(* Logix 5000 project; controller Soda_Pop_Machine 5069-L306ERM rev 38.11; software revision 38.02 *)

TASK MainTask (continuous, watchdog 500 ms) : MainProgram

MODULES
   Local : 5069-L306ERM (5069 0, rev 38.11)
       : 5069-IB16 (5069 1, rev 2.16, StandardDataDriven RPI 5 ms)
       : 5069-OB16 (5069 2, rev 3.13, StandardDataDriven RPI 5 ms)
       : 5069-IF8 (5069 3, rev 3.11, StandardDataDriven RPI 100 ms)
       : vendor 1 type 115 code 320 (5069 4, rev 2.13, StandardDataDriven RPI 80 ms)
END_MODULES

PROGRAM MainProgram   (* main routine Main *)
VAR
   Add_ice : SFC_STEP := (Status := 16#0020_0001, PauseTimer := 1, PRE := 3000);
   Add_ice_action : SFC_ACTION := (Status := 16#0020_0000, PauseTimer := 1);
   Coin : BOOL;
   Cup : STRING;
   DISPENSE : SFC_STEP := (Status := 16#0020_0001, PauseTimer := 1, PRE := 2000);
   Dispense_action : SFC_ACTION := (Status := 16#0020_0000, PauseTimer := 1);
   Drop_Cup : SFC_STEP := (Status := 16#0020_0001, PauseTimer := 1);
   Enter : BOOL;
   Finish : SFC_STEP := (Status := 16#0020_0001, PauseTimer := 1);
   Flash_lights : SFC_ACTION := (Status := 16#0020_0000, PauseTimer := 1);
   GrapeSTR : STRING := 'Grape';
   IceSTR : STRING := ' + Ice';
   INIT : SFC_STEP := (Status := 16#a820_0201, X := 1, SA := 1, DN := 1, PauseTimer := 1, T := 18659, TMax := 18659, Count := 1);
   Init_action : SFC_ACTION := (Status := 16#c020_0000, A := 1, Q := 1, PauseTimer := 1, Count := 1);
   LED_1 : ALIAS FOR Local:2:O.Pt00.Data;
   LED_2 : ALIAS FOR Local:2:O.Pt01.Data;
   LemonSTR : STRING := 'Lemon';
   Mixer_on : SFC_STEP := (Status := 16#0020_0001, PauseTimer := 1);
   Music_on : SFC_STEP := (Status := 16#0020_0001, PauseTimer := 1);
   Music_on_action : SFC_ACTION := (Status := 16#0020_0000, PauseTimer := 1);
   NullSTR : STRING;
   OrangeSTR : STRING := 'Orange';
   Pass_to_finish : BOOL;
   Pass_to_mixer : BOOL;
   Pass_to_mixer_action : SFC_ACTION := (Status := 16#0020_0000, PauseTimer := 1);
   PeachSTR : STRING := 'Peach';
   pop_type : STRING;
   Return_to_init : BOOL;
   SELECT : SFC_STEP := (Status := 16#0020_0001, PauseTimer := 1);
   Select_action : SFC_ACTION := (Status := 16#0020_0000, PauseTimer := 1);
   Socket_1 : ALIAS FOR Local:2:O.Pt02.Data;
   Socket_2 : ALIAS FOR Local:2:O.Pt03.Data;
   Switch_1 : ALIAS FOR Local:1:I.Pt00.Data;
   Switch_2 : ALIAS FOR Local:1:I.Pt01.Data;
   Switch_3 : ALIAS FOR Local:1:I.Pt02.Data;
   Switch_4 : ALIAS FOR Local:1:I.Pt03.Data;
   Switch_5 : ALIAS FOR Local:1:I.Pt04.Data;
   Switch_6 : ALIAS FOR Local:1:I.Pt05.Data;
   Wait_for_drop : BOOL;
   Wait_for_mixer : BOOL;
   Wait_for_mixer_action : SFC_ACTION := (Status := 16#0020_0000, PauseTimer := 1);
END_VAR

ROUTINE Main   (* sequential function chart *)
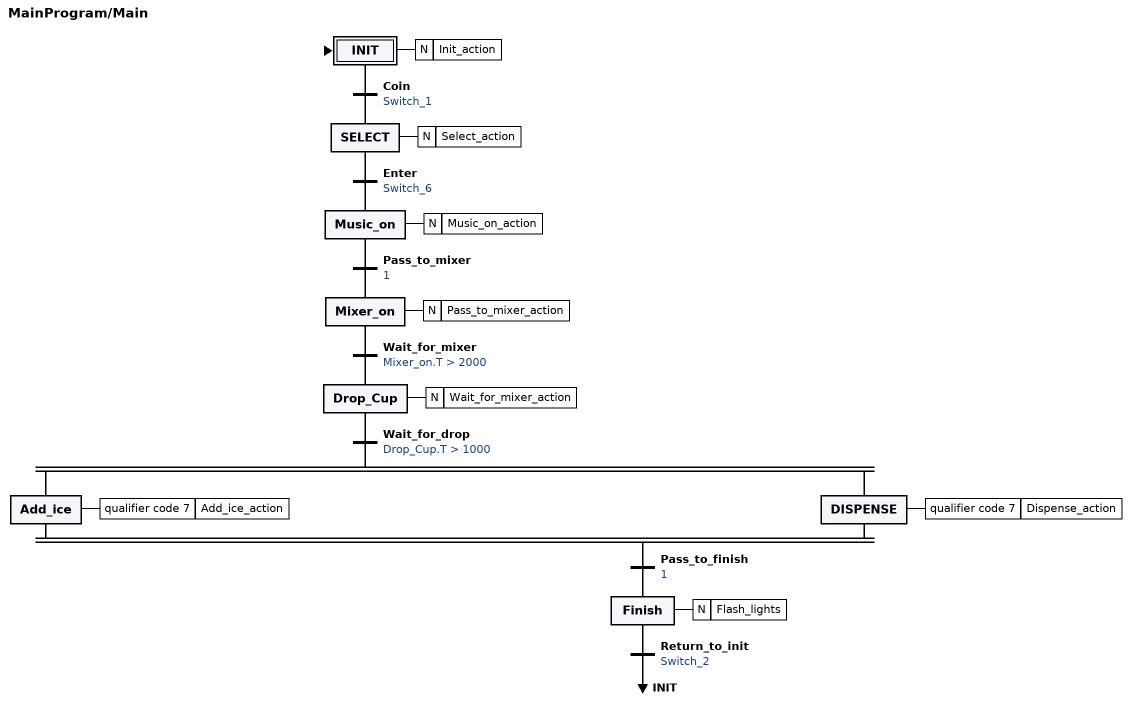
   // "add_ice"
   // step has a
   // preset wait
   // time of 3
   // seconds
   // (3000 ms)
   // "DISPENSE" step
   // has a preset wait
   // time of 2 seconds
   // (2000 ms)
   // Set initial values.
   // Turn off all LEDs
   // and sockets
   // (LEDs 3 and 4).
   // Erase cup string.
   // Select stage
   // represents the
   // customer
   // selecting a
   // options. Turn on
   // LED1 and flash
   // LED2 at 1 Hz.
   // Turn on the
   // music
   // (socket_1,
   // which is actually
   // LED3)
   // Turn on the
   // mixer (socket_2,
   // which is
   // actually LED4)
   // Wait for the
   // mixer for two
   // seconds before
   // continuing.
   // Turn off the
   // mixer. (Turn off
   // Socket_2, LED4)
   // Change the pop
   // type in the "cup"
   // string based off
   // switches 4 and
   // 5.
   // Display a
   // cascading
   // effect of LEDs
   // when finished.
   // Wait for switch
   // 2 before
   // resetting the
   // machine.
   // Wait for for the
   // selections to be
   // entered (switch
   // 6) before
   // continuing.
   INITIAL_STEP INIT:
      ACTION Init_action (N):
         LED_1 := 0;
         LED_2 := 0;
         Socket_1 := 0;
         Socket_2 := 0;
         CONCAT(NullSTR, NullSTR, Cup);
         
      END_ACTION
   END_STEP
   TRANSITION Coin FROM INIT TO SELECT
      := Switch_1
   END_TRANSITION
   STEP SELECT:
      ACTION Select_action (N):
         LED_1 := 1;
         LED_2 := ((SELECT.T / 500) MOD 2) = 0;
         
      END_ACTION
   END_STEP
   TRANSITION Enter FROM SELECT TO Music_on
      := Switch_6
   END_TRANSITION
   STEP Music_on:
      ACTION Music_on_action (N):
         Socket_1 := 1;
      END_ACTION
   END_STEP
   TRANSITION Pass_to_mixer FROM Music_on TO Mixer_on
      := 1
         
   END_TRANSITION
   STEP Mixer_on:
      ACTION Pass_to_mixer_action (N):
         Socket_2 := 1;
      END_ACTION
   END_STEP
   TRANSITION Wait_for_mixer FROM Mixer_on TO Drop_Cup
      := Mixer_on.T > 2000
         
   END_TRANSITION
   STEP Drop_Cup:
      ACTION Wait_for_mixer_action (N):
         Socket_2 := 0;
         CONCAT(NullSTR, NullSTR, Cup);
      END_ACTION
   END_STEP
   TRANSITION Wait_for_drop FROM Drop_Cup TO (DISPENSE, Add_ice)
      := Drop_Cup.T > 1000
   END_TRANSITION
   STEP Add_ice:
      ACTION Add_ice_action (qualifier code 7):
         if Switch_3 then
         	CONCAT(Cup, IceSTR, Cup);
         end_if;
      END_ACTION
   END_STEP
   STEP DISPENSE:
      ACTION Dispense_action (qualifier code 7):
         pop_type := '';
         
         
         if NOT Switch_4 AND NOT Switch_5 then
         	pop_type := OrangeSTR;
         elsif NOT Switch_4 AND Switch_5 then
         	pop_type := PeachSTR;
         elsif Switch_4 AND NOT Switch_5 then
         	pop_type := GrapeSTR;
         elsif Switch_4 AND Switch_5 then
         	pop_type := LemonSTR;
         end_if;
         
         CONCAT(Cup, pop_type, Cup);
      END_ACTION
   END_STEP
   TRANSITION Pass_to_finish FROM (Add_ice, DISPENSE) TO Finish
      := 1
         
   END_TRANSITION
   STEP Finish:
      ACTION Flash_lights (N):
         LED_1    := ((Finish.T / 50) MOD 4) = 0;
         LED_2    := ((Finish.T / 50) MOD 4) = 1;
         Socket_1 := ((Finish.T / 50) MOD 4) = 2;
         Socket_2 := ((Finish.T / 50) MOD 4) = 3;
      END_ACTION
   END_STEP
   TRANSITION Return_to_init FROM Finish TO INIT
      := Switch_2
         
   END_TRANSITION
END_ROUTINE
END_PROGRAM
